// TIA Portal V21 export
// export: Created 2026-10-12T12:46:15.8379324Z, ExportSetting WithDefaults, DisplayName Totally Integrated Automation Portal, DisplayVersion V21, DisplayName STEP 7 Professional, DisplayVersion V21, DisplayName STEP 7 Safety, DisplayVersion V21, DisplayName Tech WebApplication, DisplayVersion V21, DisplayName WinCC Basic/Comfort/Advanced, DisplayVersion V21, DisplayName WinCC Unified, DisplayVersion V21
Screen "ALARMS"  800x480, Number=3, Template=MAIN
  ScreenLayer 
    TextField "Template_Text field_2" at 372,62 size 84x27  Text="ALARMS"
